// SIMATIC S7-200 project (STEP 7-Micro/WIN), CPU 224XP CN REL 02.01

SYMBOL_TABLE ????1
C_1              VD100
C_0              VD110
w_k              VD180
r_k              VD190
y_k              VD120
y_k_1            VD130
y_k_2            VD140
u_k              VD150
u_k_1            VD160
u_k_2            VD170
Aa               VD200
Bb               VD210
Cc               VD220
Dd               VD230
Ee               VD240
END_SYMBOL_TABLE

ORGANIZATION_BLOCK ???:OB1
TITLE=
BEGIN
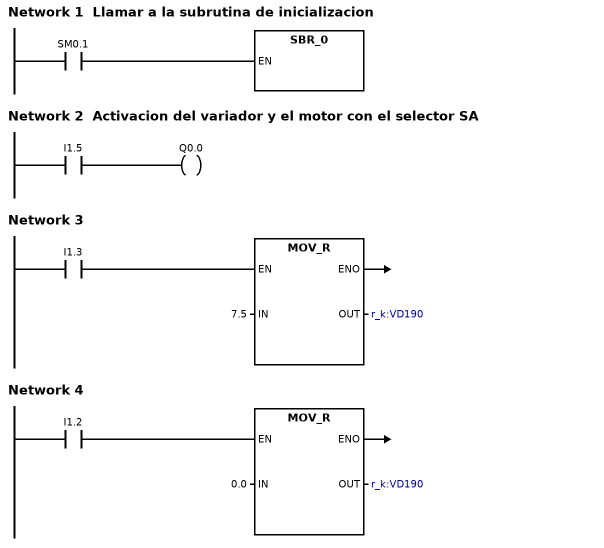
Network 1 // Llamar a la subrutina de inicializacion 
LD     SM0.1
CALL   SBR_0:SBR0
Network 2 // Activacion del variador y el motor con el selector SA
LD     I1.5
=      Q0.0
Network 3
LD     I1.3
MOVR   7.5, r_k:VD190
Network 4
LD     I1.2
MOVR   0.0, r_k:VD190
END_ORGANIZATION_BLOCK

SUBROUTINE_BLOCK SBR_0:SBR0
TITLE=
BEGIN
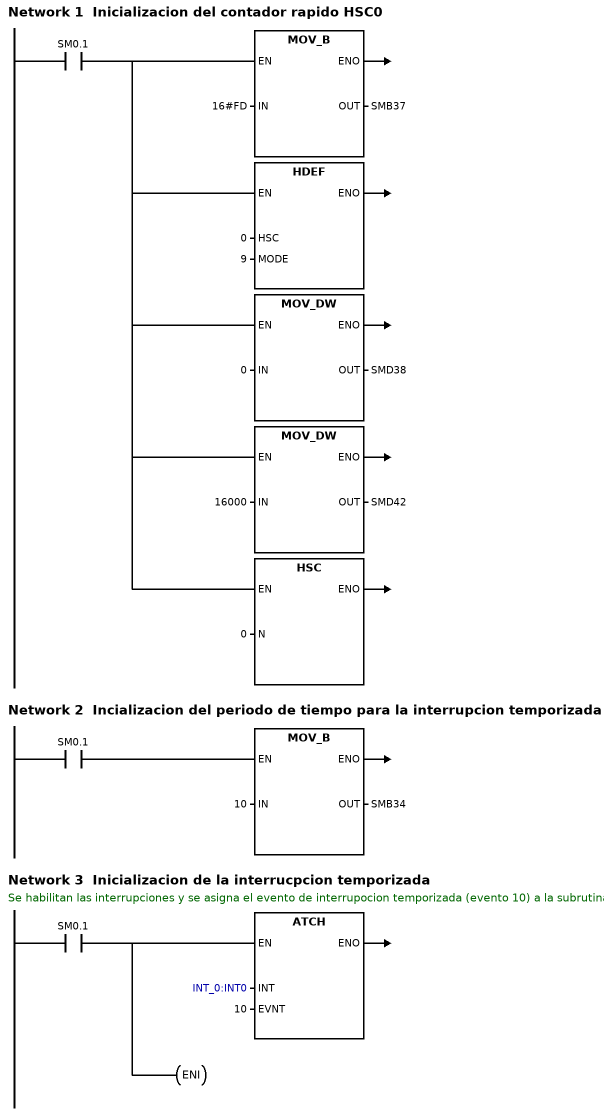
Network 1 // Inicializacion del contador rapido HSC0
LD     SM0.1
MOVB   16#FD, SMB37
HDEF   0, 9
MOVD   0, SMD38
MOVD   16000, SMD42
HSC    0
Network 2 // Incializacion del periodo de tiempo para la interrupcion temporizada
LD     SM0.1
MOVB   10, SMB34
Network 3 // Inicializacion de la interrucpcion temporizada
// Se habilitan las interrupciones y se asigna el evento de interrupocion temporizada (evento 10) a la subrutina de interrupcion INT_0
LD     SM0.1
ATCH   INT_0:INT0, 10
ENI
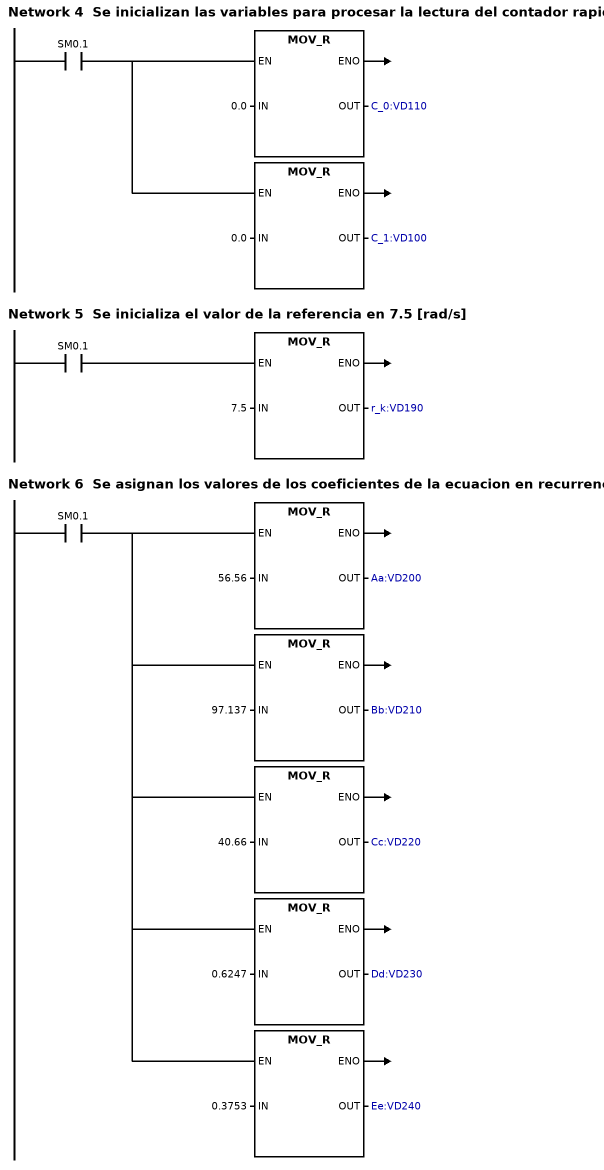
Network 4 // Se inicializan las variables para procesar la lectura del contador rapido HSC0
LD     SM0.1
MOVR   0.0, C_0:VD110
MOVR   0.0, C_1:VD100
Network 5 // Se inicializa el valor de la referencia en 7.5 [rad/s]
LD     SM0.1
MOVR   7.5, r_k:VD190
Network 6 // Se asignan los valores de los coeficientes de la ecuacion en recurrencia
LD     SM0.1
MOVR   56.56, Aa:VD200
MOVR   97.137, Bb:VD210
MOVR   40.66, Cc:VD220
MOVR   0.6247, Dd:VD230
MOVR   0.3753, Ee:VD240
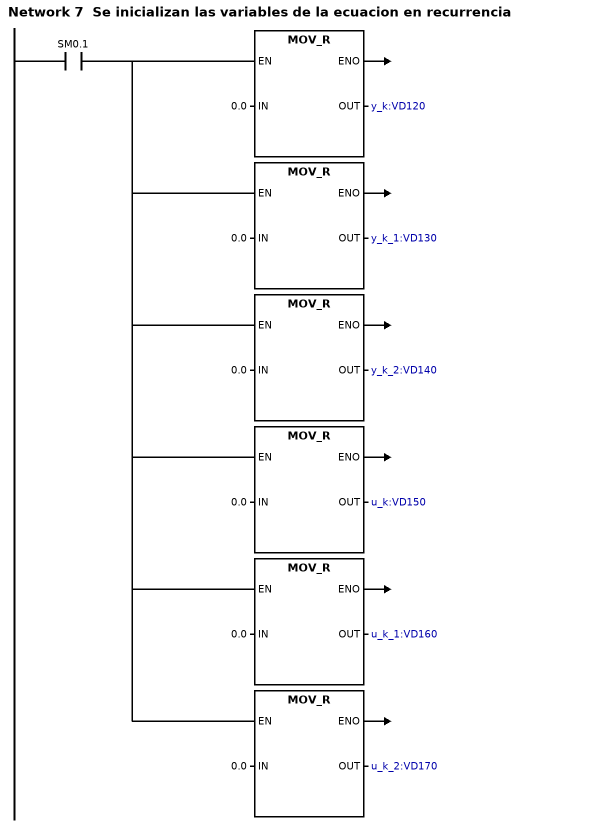
Network 7 // Se inicializan las variables de la ecuacion en recurrencia
LD     SM0.1
MOVR   0.0, y_k:VD120
MOVR   0.0, y_k_1:VD130
MOVR   0.0, y_k_2:VD140
MOVR   0.0, u_k:VD150
MOVR   0.0, u_k_1:VD160
MOVR   0.0, u_k_2:VD170
END_SUBROUTINE_BLOCK

INTERRUPT_BLOCK INT_0:INT0
TITLE=
BEGIN
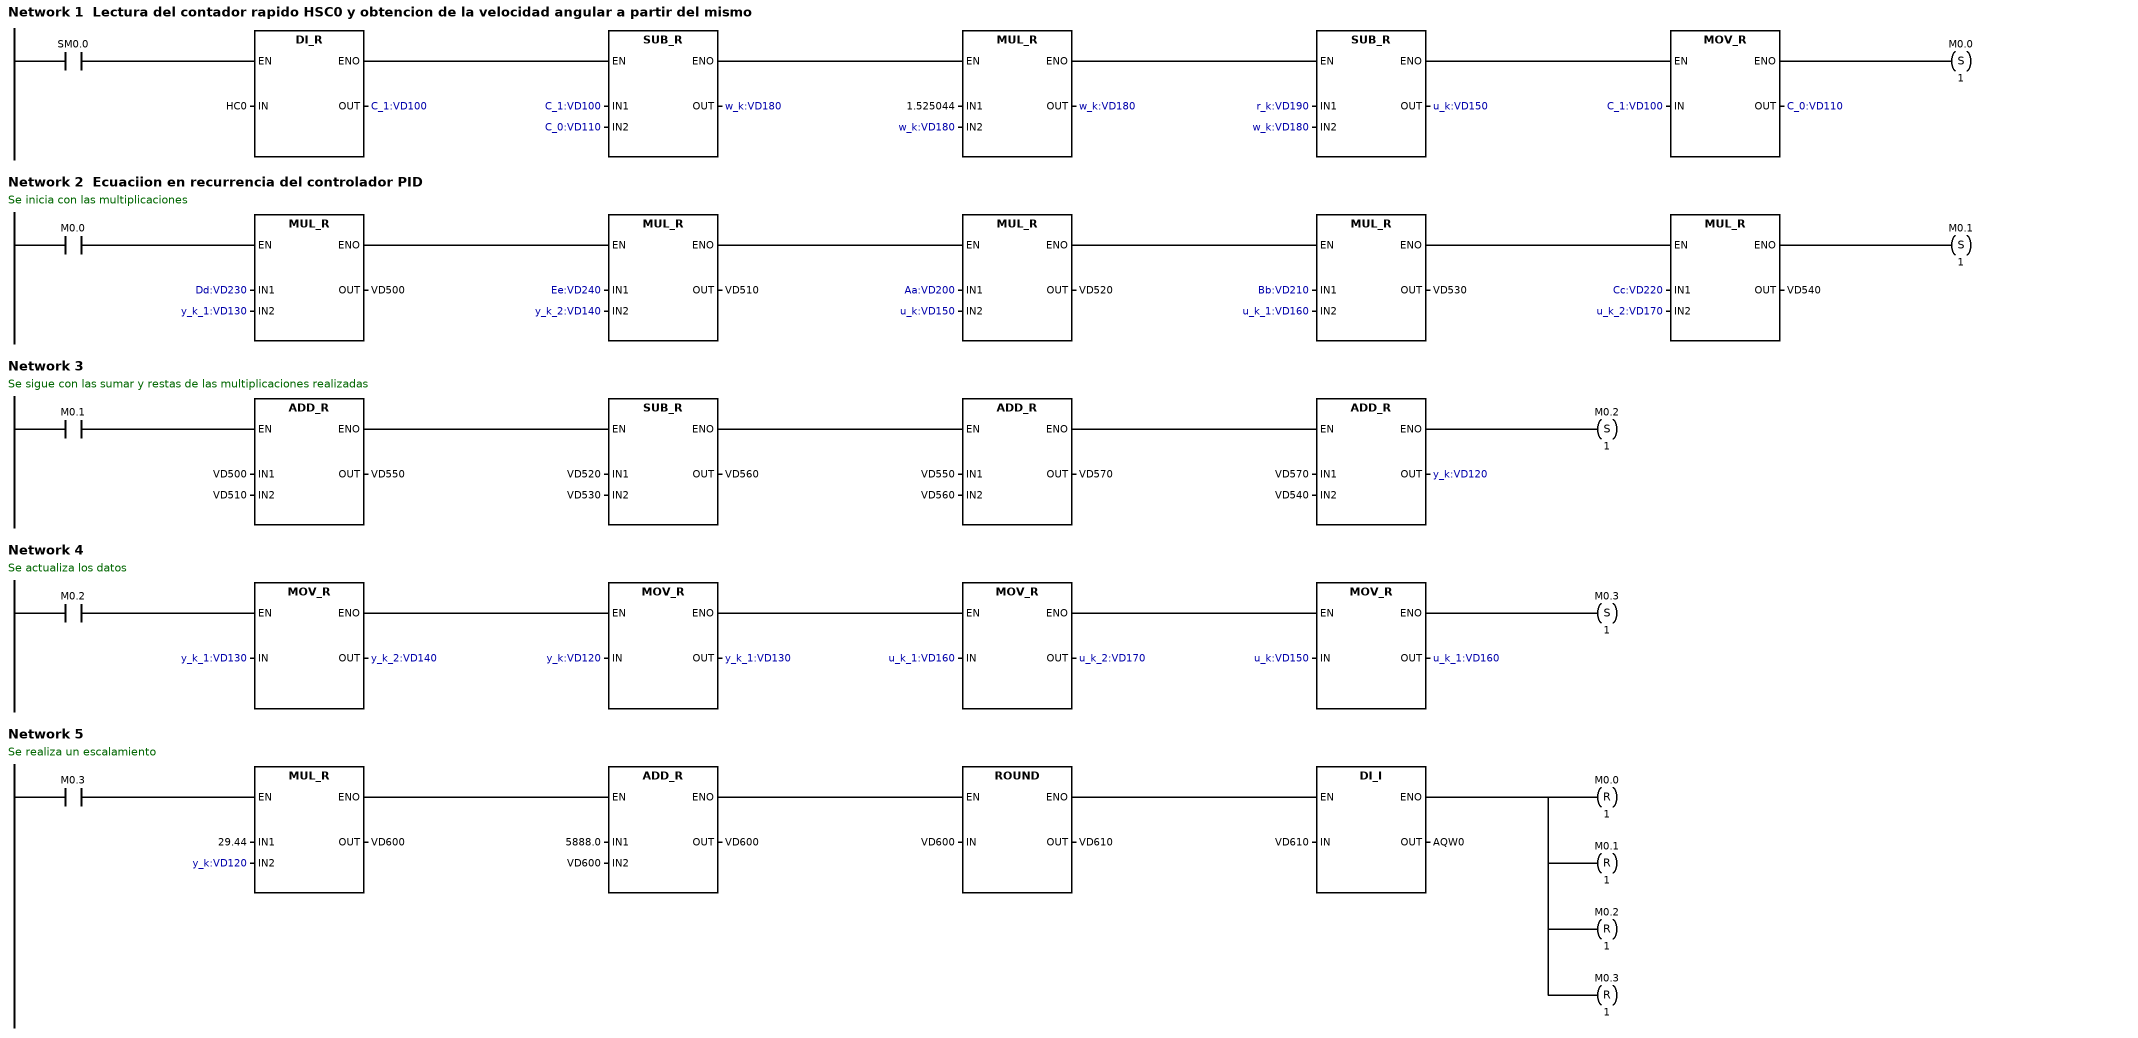
Network 1 // Lectura del contador rapido HSC0 y obtencion de la velocidad angular a partir del mismo
LD     SM0.0
DTR    HC0, C_1:VD100
AENO
MOVR   C_1:VD100, w_k:VD180
AENO
-R     C_0:VD110, w_k:VD180
AENO
*R     1.525044, w_k:VD180
AENO
MOVR   r_k:VD190, u_k:VD150
AENO
-R     w_k:VD180, u_k:VD150
AENO
MOVR   C_1:VD100, C_0:VD110
AENO
S      M0.0, 1
Network 2 // Ecuaciion en recurrencia del controlador PID
// Se inicia con las multiplicaciones
LD     M0.0
MOVR   Dd:VD230, VD500
AENO
*R     y_k_1:VD130, VD500
AENO
MOVR   Ee:VD240, VD510
AENO
*R     y_k_2:VD140, VD510
AENO
MOVR   Aa:VD200, VD520
AENO
*R     u_k:VD150, VD520
AENO
MOVR   Bb:VD210, VD530
AENO
*R     u_k_1:VD160, VD530
AENO
MOVR   Cc:VD220, VD540
AENO
*R     u_k_2:VD170, VD540
AENO
S      M0.1, 1
Network 3
// Se sigue con las sumar y restas de las multiplicaciones realizadas
LD     M0.1
MOVR   VD500, VD550
AENO
+R     VD510, VD550
AENO
MOVR   VD520, VD560
AENO
-R     VD530, VD560
AENO
MOVR   VD550, VD570
AENO
+R     VD560, VD570
AENO
MOVR   VD570, y_k:VD120
AENO
+R     VD540, y_k:VD120
AENO
S      M0.2, 1
Network 4
// Se actualiza los datos
LD     M0.2
MOVR   y_k_1:VD130, y_k_2:VD140
AENO
MOVR   y_k:VD120, y_k_1:VD130
AENO
MOVR   u_k_1:VD160, u_k_2:VD170
AENO
MOVR   u_k:VD150, u_k_1:VD160
AENO
S      M0.3, 1
Network 5
// Se realiza un escalamiento
LD     M0.3
MOVR   29.44, VD600
AENO
*R     y_k:VD120, VD600
AENO
+R     5888.0, VD600
AENO
ROUND  VD600, VD610
AENO
DTI    VD610, AQW0
AENO
R      M0.0, 1
R      M0.1, 1
R      M0.2, 1
R      M0.3, 1
END_INTERRUPT_BLOCK
